Fanuc KAREL source: kc00022.KL

-- PROVISIONAL review KL for V1013-1; original PC SHA256 3be506ab7f787f939a253f2cc9c161702d9aec00d217350d3a88be8c4c254ceb
-- Incomplete behavior may be omitted. Consult companion uncertainty JSON. Do not deploy.
PROGRAM KC00022
%NOLOCKGROUP
BEGIN
  -- UNRESOLVED_PC offsets 5-22; opcodes 3F,75
  -- UNRESOLVED_PC offsets 27-45; opcodes 27,22,2A,22,31
  -- UNRESOLVED_PC offsets 50-54; opcodes 7F
END KC00022
